{region 'Documentation'}
(*!
<summary>Real Event Buffer with command-order observations; BeginObservation excludes setup calls.</summary>
*)
{endregion}
FUNCTION_BLOCK BufferCommandProbe EXTENDS EventBuffer
VAR
    FOperationCount : UINT;
    FResetOrder : UINT;
    FResetCount : UINT;
    FDeleteCount : UINT;
END_VAR

{region 'Documentation'}
(*!
<summary>Clears only test observations, not buffer contents or reservations.</summary>
*)
{endregion}
METHOD PUBLIC BeginObservation
FOperationCount := 0;
FResetOrder := 0;
FResetCount := 0;
FDeleteCount := 0;
END_METHOD

{region 'Documentation'}
(*!
<summary>Recorded DeleteCount for command-order verification.</summary>
*)
{endregion}
{attribute 'monitoring' := 'call'}
PROPERTY PUBLIC DeleteCount : UINT //! Recorded DeleteCount for command-order verification.
GET
DeleteCount := FDeleteCount;
END_GET
END_PROPERTY

{region 'Documentation'}
(*!
<summary>Counts nonzero delete commands, then delegates unchanged to the real buffer.</summary>
*)
{endregion}
METHOD PUBLIC ProcessDeleteRequest
VAR_IN_OUT
    SequenceId : UDINT; //! Pending delete watermark passed through to the inherited consumer, which clears the request.
END_VAR
IF SequenceId <> 0 THEN
    FDeleteCount := FDeleteCount + 1;
END_IF;
SUPER^.ProcessDeleteRequest(SequenceId := SequenceId);
END_METHOD

{region 'Documentation'}
(*!
<summary>Records a Suite release attempt in the same order domain as Reset.</summary>
*)
{endregion}
METHOD PUBLIC RecordRelease : UINT //! Incremented operation sequence number shared with buffer Reset observations.
FOperationCount := FOperationCount + 1;
RecordRelease := FOperationCount;
END_METHOD

{region 'Documentation'}
(*!
<summary>Records entry, then executes the unchanged real hard reset.</summary>
*)
{endregion}
METHOD PUBLIC Reset
FOperationCount := FOperationCount + 1;
FResetOrder := FOperationCount;
FResetCount := FResetCount + 1;
SUPER^.Reset();
END_METHOD

{region 'Documentation'}
(*!
<summary>Recorded ResetCount for command-order verification.</summary>
*)
{endregion}
{attribute 'monitoring' := 'call'}
PROPERTY PUBLIC ResetCount : UINT //! Recorded ResetCount for command-order verification.
GET
ResetCount := FResetCount;
END_GET
END_PROPERTY

{region 'Documentation'}
(*!
<summary>Recorded ResetOrder for command-order verification.</summary>
*)
{endregion}
{attribute 'monitoring' := 'call'}
PROPERTY PUBLIC ResetOrder : UINT //! Recorded ResetOrder for command-order verification.
GET
ResetOrder := FResetOrder;
END_GET
END_PROPERTY

END_FUNCTION_BLOCK

(* stored: Version 1.1.0.1
   POU BufferCommandProbe: Id {4a1a79a1-4b11-45aa-896b-1313883b2c95}, SpecialFunc None
   Method BeginObservation: Id {fbe11983-8805-4bb8-892c-bfb625539b5e}
   Property DeleteCount: Id {23c1c274-87bb-49dd-9a9f-b4891a899c0e}
   Get Get: Id {8c566c29-a49e-4c4a-8696-bf97c5b862bb}
   Method ProcessDeleteRequest: Id {fc339740-4b67-4eb7-98f4-2dc09923c70d}
   Method RecordRelease: Id {1fb633e2-7c21-409f-946e-c261f3a29b83}
   Method Reset: Id {231d6610-4709-46a1-b8f5-9295f236b307}
   Property ResetCount: Id {1bf08b79-2a19-445b-b79c-7814150f706c}
   Get Get: Id {54db9886-8b32-4a5e-a0dd-f8a0705b43eb}
   Property ResetOrder: Id {4bb794e9-ee04-4b3f-bafb-6bf0d57adb15}
   Get Get: Id {3ac8839a-b67f-41a6-91d0-5d8125a1a055} *)
